TestServices.ReportAssertionFailure(
	testCase := _TestCase,
	message := _Message,
	sourceClassName := ClassName,
	defaultMessage := diagnostic
);
END_METHOD

END_FUNCTION_BLOCK

// ---- Assertions/TypedContexts/PointerAssertionContext.TcPOU
(*
SPDX-FileCopyrightText: © 2026 Oleksandr Tiutyk <trofimich@gmail.com>
SPDX-License-Identifier: MIT
License: https://opensource.org/license/mit
*)

(*!
<summary>Provides fluent assertions on a copied PVOID value.</summary>
<description>
Copies actual into persistent instance storage before the entry method returns; literals and expression
results therefore remain valid throughout the immediate chain. Owns no heap allocation or pointed-to resource.
The message prefixes every failure until the next preparation. Finish one chain before starting another on
the owning Assertions provider. Use only from the owning test callback on one task, without reentry.
Obtain this context from the owning provider; direct unprepared use is unsupported.
Expected arguments use the declared IEC type; ordinary compiler conversions happen before comparison.
This context does not depend on another assertion context.
Object metadata is available before preparation; inherited equality compares instance identity.
Copies the pointer value into a POINTER TO BYTE slot and never dereferences its target.
Equality compares addresses without generic conversion. Failed comparisons format the numeric addresses.
For interfaces and references, use ThatBool with the explicit null or validity predicate.
</description>
*)

{attribute 'no_explicit_call' := 'do not call this function block directly'}
FUNCTION_BLOCK PointerAssertionContext EXTENDS TOF_Core.Object
VAR_STAT
	{attribute 'hide'}
	_ClassName : STRING := __POUNAME();
END_VAR
VAR
	_Actual : POINTER TO BYTE;
	_TestCase : ITestCase;
	_Message : WSTRING(255);
END_VAR

(*!
<summary>Provides the implementation class name.</summary>
<description>
Borrowed read-only reference to compiler-initialized storage, valid throughout the instance lifetime.
Do not modify the returned reference; no ownership is transferred.
</description>
*)
{attribute 'monitoring' := 'call'}
PROPERTY ClassName : REFERENCE TO STRING
GET
ClassName REF= _ClassName;
END_GET
END_PROPERTY

(*!
<summary>Asserts that the copied pointer value is non-null.</summary>
<description>
Records failure without interrupting the callback; preserves the chain message.
</description>
*)
METHOD FINAL IsNotNull : REFERENCE TO PointerAssertionContext
IF _Actual = TOF_Core.Memory.NULL_ADDRESS THEN
	TestServices.ReportAssertionFailure(
		testCase := _TestCase,
		message := _Message,
		sourceClassName := ClassName,
		defaultMessage := "Expected: non-null object/pointer, but was null (0)"
	);
END_IF

IsNotNull REF= THIS^;
END_METHOD

(*!
<summary>Asserts that the copied pointer value is null.</summary>
<description>
Records failure without interrupting the callback; preserves the chain message.
</description>
*)
METHOD FINAL IsNull : REFERENCE TO PointerAssertionContext
IF _Actual <> TOF_Core.Memory.NULL_ADDRESS THEN
	TestServices.ReportAssertionFailure(
		testCase := _TestCase,
		message := _Message,
		sourceClassName := ClassName,
		defaultMessage := "Expected: null (0), but was non-zero address"
	);
END_IF

IsNull REF= THIS^;
END_METHOD

(*!
<summary>Provides the library namespace.</summary>
<description>
Borrowed read-only reference to the compiler-initialized namespace, valid throughout the instance lifetime.
Do not modify the returned reference; no ownership is transferred.
</description>
*)
{attribute 'monitoring' := 'call'}
PROPERTY NamespaceName : REFERENCE TO STRING
GET
NamespaceName REF= CurrentNamespace.Name;
END_GET
END_PROPERTY

(*!
<summary>Asserts inequality with the expected value.</summary>
<description>
Records failure without interrupting the callback; preserves the message for the rest of the chain.
</description>
<param name="expected">Expected value converted by the compiler to PVOID.</param>
*)
METHOD FINAL NotToBe : REFERENCE TO PointerAssertionContext
VAR_INPUT
	expected : PVOID;
END_VAR
IF _Actual = expected THEN
	failComparison(
		expected := expected,
		expectation := "Expected value not to be: "
	);
END_IF

NotToBe REF= THIS^;
END_METHOD

(*!
<summary>Copies the actual operand and replaces the chain-wide message.</summary>
<description>
Called by the owning Assertions provider after it verifies the running test case.
No pointer to this method's input storage is retained. The receiver is borrowed until the next preparation;
the owning provider keeps it alive throughout the immediate chain.
</description>
<param name="actual">Value copied into this context.</param>
<param name="testCase">Borrowed failure receiver for the immediate chain.</param>
<param name="message">Copied diagnostic prefix, including empty to clear the previous prefix.</param>
*)
METHOD INTERNAL FINAL Prepare
VAR_INPUT
	actual : PVOID;
	testCase : ITestCase;
	message : WSTRING(255);
END_VAR
_Actual := actual;
_TestCase := testCase;
_Message := message;
END_METHOD

(*!
<summary>Reports the byte size of this concrete instance.</summary>
<description>
Includes inline fields and nested instances, but excludes separately allocated payloads.
Obtaining the size does not transfer ownership or validate an arbitrary address.
</description>
*)
{attribute 'monitoring' := 'call'}
PROPERTY SelfSize : ULINT
GET
SelfSize := XSIZEOF(THIS^);
END_GET
END_PROPERTY

(*!
<summary>Asserts equality with the expected value.</summary>
<description>
Records failure without interrupting the callback; preserves the message for the rest of the chain.
</description>
<param name="expected">Expected value converted by the compiler to PVOID.</param>
*)
METHOD FINAL ToBe : REFERENCE TO PointerAssertionContext
VAR_INPUT
	expected : PVOID;
END_VAR
IF _Actual <> expected THEN
	failComparison(
		expected := expected,
		expectation := "Expected: "
	);
END_IF

ToBe REF= THIS^;
END_METHOD

(*!
<summary>Formats a failed typed predicate and reports it with the chain message.</summary>
<description>
Does not change operands or chain state. The receiver retains its first failure. Reporting exceptions
propagate to the enclosing test callback handler; an unprepared receiver is a configuration error.
</description>
<param name="expected">Typed expected operand used only for this diagnostic.</param>
<param name="expectation">Prefix identifying the failed predicate.</param>
*)
METHOD PRIVATE failComparison
VAR_INPUT
	expected : PVOID;
	expectation : WSTRING(40);
END_VAR
VAR
	actualText : WSTRING(255);
	expectedText : WSTRING(255);
	diagnostic : TOF_Core.ERROR_MESSAGE;
END_VAR
actualText := TO_WSTRING(TO_ULINT(_Actual));
expectedText := TO_WSTRING(TO_ULINT(expected));

diagnostic := TOF_Core.WideStrings.Concat255(
	expectation,
	expectedText,
	", but was: ",
	actualText
);

TestServices.ReportAssertionFailure(
	testCase := _TestCase,
	message := _Message,
	sourceClassName := ClassName,
	defaultMessage := diagnostic
);
END_METHOD

END_FUNCTION_BLOCK

// ---- TestElements/Groups/TestGroup.TcPOU
(*
SPDX-FileCopyrightText: © 2026 Oleksandr Tiutyk <trofimich@gmail.com>
SPDX-License-Identifier: MIT
License: https://opensource.org/license/mit
*)

(*!
<summary>Executes the fixed child array provided by a concrete group.</summary>
<description>
Descendants own persistent tests, nested groups and interface-array storage. Children returns the same valid
array throughout the group lifetime; callers must not modify its contents through the reference. Each child
is non-null, occurs once and has this group as its constructor-assigned Parent. Parent chains are acyclic.
All objects outlive the tree; no allocation ownership is transferred. Zero children form an empty group.
Reset validates the child reference, slots and parent chain once at the start of each run. Missing
array storage raises DataMemberNotSpecifiedException; null slots do likewise with an indexed member name.
Duplicates, a mismatched parent or a parent cycle raise StandardException before any direct child is called.
A descendant's validation or callback can still fail after earlier siblings have reset; no rollback is promised.
Execute drives one current child once and counts it once when finished. Groups add no synthetic test results
and have no scenario setup or teardown hooks. Use the entire tree in one task without reentry.
Do not mutate the child array or parent associations during the lifetime of the tree, or copy instances by value.
</description>
*)

{attribute 'no_explicit_call' := 'do not call this function block directly'}
FUNCTION_BLOCK ABSTRACT TestGroup
VAR_GENERIC CONSTANT
	//! <summary>Exact number of direct child slots; zero produces an empty array.</summary>
	{attribute 'hide'} 
	_ChildCount : TOF_Core.INT_LENGTH := 0;
END_VAR
EXTENDS TestElement IMPLEMENTS IParentTestElement
VAR
	{attribute 'hide'} 
	_CurrentChildIndex : TOF_Core.INT_LENGTH;
	
	{attribute 'hide'} 
	_TestCount : TOF_Core.DINT_LENGTH;
END_VAR

(*!
<summary>Reports the generic number of direct children.</summary>
*)

{attribute 'monitoring' := 'call'}
PROPERTY FINAL ChildCount : TOF_Core.INT_LENGTH
GET
ChildCount := _ChildCount;
END_GET
END_PROPERTY

(*!
<summary>Borrows the concrete group's persistent fixed array of tests and nested groups.</summary>
<description>
Return the same valid storage and unchanged child list for the group lifetime, including an empty array
when the generic count is zero. The getter must have no side effects. Callers may only read the reference.
Children are borrowed; each has this group as its fixed Parent and remains alive while the tree is used.
The base constructor never reads this property. Reset validates it before execution starts.
</description>
*)
{attribute 'monitoring' := 'call'}
PROPERTY ABSTRACT Children : REFERENCE TO ARRAY [0.._ChildCount - 1] OF ITestElement
GET
END_GET
END_PROPERTY

(*!
<summary>Advances one child of the validated fixed composition and counts it once on completion.</summary>
<description>
Requires a successful Reset before the first execution and every subsequent run, including after a failed Reset.
Uses the concrete group's Children reference without repeating topology validation.
External exceptions propagate to the runner and abort the run.
Neither Reset nor Execute changes parent associations.
</description>
*)
METHOD FINAL Execute
VAR
	childElements : REFERENCE TO ARRAY [0.._ChildCount - 1] OF ITestElement;
END_VAR
IF IsFinished THEN
	RETURN;
END_IF

childElements REF= THIS^.Children;

_State := TEST_ELEMENT_STATE.RUNNING;
_Duration := _Duration + TOF_Core.System.GetTaskCycleTime();

IF _CurrentChildIndex < _ChildCount THEN
	childElements[_CurrentChildIndex].Execute();

	IF childElements[_CurrentChildIndex].IsFinished THEN
		_PassedCount := _PassedCount + childElements[_CurrentChildIndex].PassedCount;
		_FailedCount := _FailedCount + childElements[_CurrentChildIndex].FailedCount;
		_SkippedCount := _SkippedCount + childElements[_CurrentChildIndex].SkippedCount;
		_CurrentChildIndex := _CurrentChildIndex + 1;
	END_IF

END_IF

IF _CurrentChildIndex >= _ChildCount THEN
	_State := TEST_ELEMENT_STATE.COMPLETED;
	_Reporter := 0;
END_IF
END_METHOD

(*!
<summary>Borrows one direct child in fixed execution order without changing the tree.</summary>
<description>
Checks storage before the index, including before the first Reset and after a failed Reset.
Missing storage or a null selected slot raises DataMemberNotSpecifiedException; an index outside
zero through ChildCount minus one raises ArgumentOutOfRangeException. No child callback is invoked.
The returned interface is borrowed for the child's lifetime. Use from the owning task without reentry;
this method does not repeat complete topology validation or authorize changes to the composition.
</description>
<param name="index">Zero-based position in the fixed direct-child array.</param>
*)
METHOD FINAL GetChildByIndex : ITestElement
VAR_INPUT
	index : TOF_Core.INT_LENGTH;
END_VAR
IF NOT __ISVALIDREF(Children) THEN
	TOF_Core.Exceptions.ThrowDataMemberNotSpecified(
		sourceNamespaceName := NamespaceName,
		sourceClassName := ClassName,
		sourcePOUName := __POUNAME(),
		sourcePosition := __POSITION(),
		dataMemberName := 'Children'
	);
END_IF

IF index < TOF_Core.SignedInt16.ZERO OR_ELSE index >= _ChildCount THEN
	TOF_Core.Exceptions.ThrowArgumentOutOfRange(
		sourceNamespaceName := NamespaceName,
		sourceClassName := ClassName,
		sourcePOUName := __POUNAME(),
		sourcePosition := __POSITION(),
		argumentName := 'index',
		argumentValue := index
	);
END_IF

IF Children[index] = 0 THEN
	TOF_Core.Exceptions.ThrowDataMemberNotSpecified(
		sourceNamespaceName := NamespaceName,
		sourceClassName := ClassName,
		sourcePOUName := __POUNAME(),
		sourcePosition := __POSITION(),
		dataMemberName := TOF_Core.Strings.Concat255('Children[', TO_STRING(index), ']')
	);
END_IF

GetChildByIndex := Children[index];
END_METHOD

//! <summary>Sums the leaf counts of the group's direct children.</summary>
METHOD PRIVATE getTestCount : TOF_Core.DINT_LENGTH
VAR
	// An empty group gives the FOR loop an upper bound of -1.
	i : INT;
END_VAR
IF NOT __ISVALIDREF(Children) THEN
	RETURN;
END_IF

FOR i := 0 TO _ChildCount - 1 DO
	getTestCount := getTestCount + Children[i].TestCount;
END_FOR
END_METHOD

(*!
<summary>Clears observations and recursively resets descendant-specific state.</summary>
<description>
Does not run teardown or release user resources. Call only at the lifecycle boundaries in ITestElement.
The reporter is borrowed until completion; no locks or cross-task transfer are provided.
Validation or a child Reset exception propagates and can leave a partially reset tree; the runner aborts startup.
</description>
*)
METHOD FINAL Reset
VAR_INPUT
	reporter : ITestReporter;
END_VAR
VAR
	self : ITestElement;
	slowAncestor : ITestElement;
	fastAncestor : ITestElement;
	childParent : ITestElement;

	i : INT;
	j : INT;
	
	errorMessage : TOF_Core.ERROR_MESSAGE;
END_VAR
SUPER^.Reset(reporter := reporter);

IF NOT __ISVALIDREF(Children) THEN
	TOF_Core.Exceptions.ThrowDataMemberNotSpecified(
		sourceNamespaceName := NamespaceName,
		sourceClassName := ClassName,
		sourcePOUName := __POUNAME(),
		sourcePosition := __POSITION(),
		dataMemberName := 'Children'
	);
END_IF

self := THIS^;
slowAncestor := self;
fastAncestor := self;

// Traverse the fixed parent chain at two speeds to detect cycles without allocation or recursion.
WHILE fastAncestor <> 0 DO
	fastAncestor := fastAncestor.Parent;

	IF fastAncestor = 0 THEN
		EXIT;
	END_IF

	fastAncestor := fastAncestor.Parent;
	slowAncestor := slowAncestor.Parent;

	IF fastAncestor <> 0 AND_THEN fastAncestor = slowAncestor THEN
		TOF_Core.Exceptions.ThrowStandard(
			sourceNamespaceName := NamespaceName,
			sourceClassName := ClassName,
			sourcePOUName := __POUNAME(),
			sourcePosition := __POSITION(),
			message := "The assigned parent chain contains a cycle"
		);
	END_IF
END_WHILE

FOR i := 0 TO _ChildCount - 1 DO
	IF Children[i] = 0 THEN
		TOF_Core.Exceptions.ThrowDataMemberNotSpecified(
			sourceNamespaceName := NamespaceName,
			sourceClassName := ClassName,
			sourcePOUName := __POUNAME(),
			sourcePosition := __POSITION(),
			dataMemberName := TOF_Core.Strings.Concat255('Children[', TO_STRING(i), ']')
		);
	END_IF

	childParent := Children[i].Parent;

	IF childParent <> self THEN
		errorMessage := TOF_Core.WideStrings.Concat255("A child '", Children[i].Name, "' has a different constructor-assigned parent"); 
		
		TOF_Core.Exceptions.ThrowStandard(
			sourceNamespaceName := NamespaceName,
			sourceClassName := ClassName,
			sourcePOUName := __POUNAME(),
			sourcePosition := __POSITION(),
			message := errorMessage
		);
	END_IF

	FOR j := 0 TO i - 1 DO
		IF Children[i] = Children[j] THEN
			errorMessage := TOF_Core.WideStrings.Concat255("A child '", Children[i].Name, "' occupies more than one slot"); 
			
			TOF_Core.Exceptions.ThrowStandard(
				sourceNamespaceName := NamespaceName,
				sourceClassName := ClassName,
				sourcePOUName := __POUNAME(),
				sourcePosition := __POSITION(),
				message := errorMessage
			);
		END_IF
	END_FOR
END_FOR

_CurrentChildIndex := 0;

FOR i := 0 TO _ChildCount - 1 DO
	Children[i].Reset(reporter := _Reporter);
END_FOR
END_METHOD

(*!
<summary>Sums the configured leaf counts of the direct children.</summary>
<description>
Requires a valid, acyclic subtree. Traverses nested groups through their getters using the current task stack.
An empty group returns zero. Missing child storage or a null slot in a nonempty group raises
DataMemberNotSpecifiedException. Child getter exceptions propagate and the tree state is unchanged.
</description>
*)
{attribute 'monitoring' := 'call'}
PROPERTY FINAL TestCount : TOF_Core.DINT_LENGTH
GET
IF _TestCount = 0 THEN
	_TestCount := getTestCount();
END_IF

TestCount := _TestCount;
END_GET
END_PROPERTY

END_FUNCTION_BLOCK

// ---- Reporting/AdsLogReporter.TcPOU
(*
SPDX-FileCopyrightText: © 2026 Oleksandr Tiutyk <trofimich@gmail.com>
SPDX-License-Identifier: MIT
License: https://opensource.org/license/mit
*)

(*!
<summary>Writes run summaries and leaf failures to the ADS log.</summary>
<description>
Use in one task without reentry. The ADS backend has no established concurrent-call guarantee, even for
separate reporter instances. For multiple tasks use per-task in-memory reports or a synchronized backend.
Each callback submits at most one record. The ADS completion record includes counts and the first failed leaf name.
LastRunSummary includes the first failed leaf name and a bounded
version of its diagnostic. The summary and failed log writes are observable after the run. A failed
write does not change the test outcome. Individual ADS failure records are capped at 200 wide characters.
ReportRunStart clears all observations before attempting the start message.
</description>
*)

{attribute 'no_explicit_call' := 'do not call this function block directly'}
FUNCTION_BLOCK AdsLogReporter EXTENDS TOF_Core.Object IMPLEMENTS ITestReporter
VAR_STAT
	_ClassName : STRING := __POUNAME();
END_VAR
VAR
	_AdsLogger : TOF_Core.AdsLogger;
	_FirstFailureName : WSTRING;
	_FirstFailureDiagnostic : WSTRING(255);
	_LastRunSummary : TOF_Core.ERROR_MESSAGE;
	_FailedLogWriteCount : UDINT;
	_LastLogFailureMessage : TOF_Core.ERROR_MESSAGE;
END_VAR

(*!
<summary>Provides the implementation class name.</summary>
*)
{attribute 'monitoring' := 'call'}
PROPERTY ClassName : REFERENCE TO STRING
GET
ClassName REF= _ClassName;
END_GET
END_PROPERTY

(*!
<summary>Counts start, result and summary writes for which TryLogMessage returned FALSE.</summary>
<description>The count resets at ReportRunStart. A successful write does not confirm display in XAE.</description>
*)
{attribute 'monitoring' := 'call'}
PROPERTY FailedLogWriteCount : UDINT
GET
FailedLogWriteCount := _FailedLogWriteCount;
END_GET
END_PROPERTY

(*!
<summary>Borrows the last message whose ADS logger call returned FALSE.</summary>
<description>Empty until a write fails in the current run. Callers must not modify the returned storage.</description>
*)
{attribute 'monitoring' := 'call'}
PROPERTY LastLogFailureMessage : REFERENCE TO TOF_Core.ERROR_MESSAGE
GET
LastLogFailureMessage REF= _LastLogFailureMessage;
END_GET
END_PROPERTY

(*!
<summary>Borrows the summary created at ReportRunEnd regardless of its ADS write status.</summary>
<description>Empty after ReportRunStart until ReportRunEnd. Callers must not modify the returned storage.</description>
*)
{attribute 'monitoring' := 'call'}
PROPERTY LastRunSummary : REFERENCE TO TOF_Core.ERROR_MESSAGE
GET
LastRunSummary REF= _LastRunSummary;
END_GET
END_PROPERTY

(*!
<summary>Submits one ADS message and records a FALSE result from the logger.</summary>
<description>The count saturates at the largest UDINT. The copied text remains available until the next start.</description>
*)
METHOD PRIVATE logMessage
VAR_INPUT
	category : TOF_Core.LOG_CATEGORY;
END_VAR
VAR_IN_OUT CONSTANT
	message : TOF_Core.ERROR_MESSAGE;
END_VAR
IF TryWriteMessage(category := category, message := message) THEN
	RETURN;
END_IF

IF _FailedLogWriteCount < TOF_Core.UnsignedInt32.MAX_VALUE THEN
	_FailedLogWriteCount := _FailedLogWriteCount + 1;
END_IF

_LastLogFailureMessage := message;
END_METHOD

(*!
<summary>Provides the library namespace.</summary>
*)
{attribute 'monitoring' := 'call'}
PROPERTY NamespaceName : REFERENCE TO STRING
GET
NamespaceName REF= CurrentNamespace.Name;
END_GET
END_PROPERTY

(*!
<summary>Logs leaf counts and the first failed leaf name and retains its diagnostic for online inspection.</summary>
<description>The retained summary also includes a bounded first-failure diagnostic and survives a rejected ADS write.</description>
*)
METHOD ReportRunEnd
VAR_INPUT
	totalTests : TOF_Core.DINT_LENGTH;
	passedTests : TOF_Core.DINT_LENGTH;
	failedTests : TOF_Core.DINT_LENGTH;
	skippedTests : TOF_Core.DINT_LENGTH;
	duration : TIME;
END_VAR
VAR
	logSummary : WSTRING(255);
	logRecord : TOF_Core.ERROR_MESSAGE;
	summary : WSTRING(255);
END_VAR
summary := TOF_Core.WideStrings.Concat255(
	"[TOF_Testing] Finished: ", TO_WSTRING(passedTests), " passed, ",
	TO_WSTRING(failedTests), " failed, ", TO_WSTRING(skippedTests), " skipped"
);

logSummary := summary;

IF failedTests > 0 AND_THEN _FirstFailureDiagnostic <> "" THEN
	TOF_Core.WideStrings.AppendFit255(logSummary, " | First failed test: ", _FirstFailureName);
	TOF_Core.WideStrings.AppendFit255(summary, " | First failure: ", _FirstFailureDiagnostic);
END_IF

_LastRunSummary := summary;
logRecord := logSummary;
logMessage(category := TOF_Core.LOG_CATEGORY.INFORMATION, message := logRecord);
END_METHOD

(*!
<summary>Resets per-run observations and logs the number of configured leaf tests.</summary>
<description>A failed start-message write counts toward the new run.</description>
*)
METHOD ReportRunStart
VAR_INPUT
	testCount : TOF_Core.DINT_LENGTH;
END_VAR
VAR
	diagnostic : TOF_Core.ERROR_MESSAGE;
END_VAR
_FirstFailureName := "";
_FirstFailureDiagnostic := "";
_LastRunSummary := "";
_FailedLogWriteCount := 0;
_LastLogFailureMessage := "";

diagnostic := TOF_Core.WideStrings.Concat255(
	"[TOF_Testing] Starting ", TO_WSTRING(testCount), " tests"
);

logMessage(category := TOF_Core.LOG_CATEGORY.INFORMATION, message := diagnostic);
END_METHOD

(*!
<summary>Logs a failed leaf with its group path and caches the first failure for the summary.</summary>
<description>
The individual ADS record uses up to 200 wide characters to leave room below the native ADS text limit.
The retained summary includes the leaf name and the beginning of its diagnostic.
</description>
<param name="testName">Individual name bounded to 80 wide characters, matching INamed.</param>
*)
METHOD ReportTestCaseResult
VAR_INPUT
	groupPath : WSTRING(255);
	testName : WSTRING;
	outcome : TEST_OUTCOME;
	duration : TIME;
END_VAR
VAR_IN_OUT CONSTANT
	message : TOF_Core.ERROR_MESSAGE;
END_VAR
VAR
	shortDiagnostic : WSTRING(200);
	diagnostic : TOF_Core.ERROR_MESSAGE;
END_VAR
IF outcome <> TEST_OUTCOME.PASSED
	AND_THEN outcome <> TEST_OUTCOME.FAILED
	AND_THEN outcome <> TEST_OUTCOME.SKIPPED
THEN
	TOF_Core.Exceptions.ThrowArgumentValueNotSupported(
		sourceNamespaceName := NamespaceName,
		sourceClassName := ClassName,
		sourcePOUName := __POUNAME(),
		sourcePosition := __POSITION(),
		argumentName := 'outcome',
		argumentValue := outcome
	);
END_IF

IF outcome <> TEST_OUTCOME.FAILED THEN
	RETURN;
END_IF

IF _FirstFailureDiagnostic = "" THEN
	_FirstFailureName := testName;

	IF _FirstFailureName = "" THEN
		_FirstFailureName := "<unnamed>";
	END_IF

	_FirstFailureDiagnostic := TOF_Core.WideStrings.Concat255(_FirstFailureName, ": ");
	TOF_Core.WideStrings.AppendFit(targetString := _FirstFailureDiagnostic, sourceString := message);
END_IF

shortDiagnostic := "[TOF_Testing] ";

IF groupPath <> "" THEN
	TOF_Core.WideStrings.AppendFit255(shortDiagnostic, groupPath, "/");
END_IF

TOF_Core.WideStrings.AppendFit255(shortDiagnostic, testName, ": ");
TOF_Core.WideStrings.AppendFit(targetString := shortDiagnostic, sourceString := message);
diagnostic := shortDiagnostic;

logMessage(category := TOF_Core.LOG_CATEGORY.ERROR, message := diagnostic);
END_METHOD

(*!
<summary>Reports instance storage without separately allocated payloads.</summary>
*)
{attribute 'monitoring' := 'call'}
PROPERTY SelfSize : ULINT
GET
SelfSize := XSIZEOF(THIS^);
END_GET
END_PROPERTY

(*!
<summary>Submits one message to the ADS backend and reports whether the logger accepted it.</summary>
<description>
An override may replace the backend. It must return FALSE on rejection and must not raise an exception,
retry the write, or retain the borrowed message. TRUE does not confirm display in XAE.
</description>
*)
METHOD PROTECTED TryWriteMessage : BOOL
VAR_INPUT
	category : TOF_Core.LOG_CATEGORY;
END_VAR
VAR_IN_OUT CONSTANT
	message : TOF_Core.ERROR_MESSAGE;
END_VAR
TryWriteMessage := _AdsLogger.TryLogMessage(category := category, message := message);
END_METHOD

END_FUNCTION_BLOCK

// ---- Reporting/JUnitXmlReporter.TcPOU
(*
SPDX-FileCopyrightText: © 2026 Oleksandr Tiutyk <trofimich@gmail.com>
SPDX-License-Identifier: MIT
License: https://opensource.org/license/mit
*)

(*!
<summary>Builds an in-memory JUnit report with one testcase per leaf.</summary>
<description>
One flat testsuite contains all leaves; testcase classname preserves the slash-separated group path.
Wide names and diagnostics are escaped as ASCII XML character references, including surrogate pairs.
XML 1.0 disallowed control characters, isolated surrogates and U+FFFE/U+FFFF are replaced by U+FFFD;
tab, line feed and carriage return are emitted as references to preserve attribute whitespace.
Use a separate instance and buffer for each runner task without reentry. Read ContentLength bytes from
ContentAddress only after IsReady and before reset or the next run. Buffer growth invalidates old addresses.
The reporter owns its dynamic buffer; never copy it by value. Callback exceptions can leave incomplete XML.
</description>
*)

{attribute 'no_explicit_call' := 'do not call this function block directly'}
FUNCTION_BLOCK JUnitXmlReporter EXTENDS TOF_Core.Object IMPLEMENTS ITestReporter
VAR CONSTANT
	//! <summary>First and last UTF-16 high-surrogate code units; subtract the first to recover ten payload bits.</summary>
	HIGH_SURROGATE_FIRST : UDINT := 16#D800;
	//! <summary>Last UTF-16 high-surrogate code unit accepted as the first part of a pair.</summary>
	HIGH_SURROGATE_LAST : UDINT := 16#DBFF;
	//! <summary>First and last UTF-16 low-surrogate code units; subtract the first to recover ten payload bits.</summary>
	LOW_SURROGATE_FIRST : UDINT := 16#DC00;
	//! <summary>Last UTF-16 low-surrogate code unit; isolated surrogates through this value are invalid scalars.</summary>
	LOW_SURROGATE_LAST : UDINT := 16#DFFF;
	//! <summary>Base scalar value added when decoding a supplementary UTF-16 surrogate pair.</summary>
	SUPPLEMENTARY_FIRST : UDINT := 16#10000;
	//! <summary>Multiplier that moves a high surrogate's ten payload bits above the low payload.</summary>
	SURROGATE_PAYLOAD_BASE : UDINT := 1024;
	//! <summary>Printable ASCII boundaries; these scalars are emitted as bytes instead of decimal XML references.</summary>
	PRINTABLE_ASCII_FIRST : UDINT := 32;
	//! <summary>Last ASCII scalar emitted directly as a byte instead of a decimal XML reference.</summary>
	PRINTABLE_ASCII_LAST : UDINT := 126;
END_VAR
VAR_STAT
	_ClassName : STRING := __POUNAME();
END_VAR
VAR
	_Buffer : TOF_Core.StringBuilder;
	_IsReady : BOOL;
END_VAR

//! <summary>Escapes UTF-16 input and replaces isolated surrogates and forbidden XML characters.</summary>
METHOD PRIVATE appendEscapedText
VAR_IN_OUT CONSTANT
	text : WSTRING;
END_VAR
VAR
	charLength : UDINT;
	i : UDINT;
	wordPointer : POINTER TO WORD;
	codePoint : UDINT;
END_VAR
charLength := TOF_Core.WideStrings.GetLength(value := text);
wordPointer := ADR(text);

WHILE i < charLength DO
	codePoint := wordPointer[i];
	i := i + 1;

	IF codePoint >= HIGH_SURROGATE_FIRST AND_THEN codePoint <= HIGH_SURROGATE_LAST AND_THEN i < charLength
		AND_THEN wordPointer[i] >= LOW_SURROGATE_FIRST AND_THEN wordPointer[i] <= LOW_SURROGATE_LAST
	THEN
		// UTF-16 uses high D800..DBFF and low DC00..DFFF surrogates. Subtract their bases to obtain
		// ten-bit payloads; shift the high payload by ten bits and add the supplementary-plane base.
		codePoint := SUPPLEMENTARY_FIRST + (codePoint - HIGH_SURROGATE_FIRST) * SURROGATE_PAYLOAD_BASE
			+ (wordPointer[i] - LOW_SURROGATE_FIRST);
		i := i + 1;
	END_IF

	appendXmlCharacter(codePoint := codePoint);
END_WHILE
END_METHOD

(*!
<summary>Appends a scalar as printable ASCII or an XML decimal character reference.</summary>
<description>Explicitly terminates the single-byte temporary before the buffer reads it.</description>
*)
METHOD PRIVATE appendXmlCharacter
VAR_INPUT
	codePoint : UDINT;
END_VAR
VAR
	character : STRING(1);
	referenceText : STRING(255);
END_VAR
// XML 1.0 permits only TAB/LF/CR below U+0020 and excludes surrogates and U+FFFE/U+FFFF.
CASE codePoint OF
	0..8, 11, 12, 14..31, 16#D800..16#DFFF, 16#FFFE, 16#FFFF:
		_Buffer.AppendString(value := '&#65533;');
	34:
		_Buffer.AppendString(value := '&quot;');
	38:
		_Buffer.AppendString(value := '&amp;');
	39:
		_Buffer.AppendString(value := '&apos;');
	60:
		_Buffer.AppendString(value := '&lt;');
	62:
		_Buffer.AppendString(value := '&gt;');
ELSE
	IF codePoint >= PRINTABLE_ASCII_FIRST AND_THEN codePoint <= PRINTABLE_ASCII_LAST THEN
		character[0] := TO_BYTE(codePoint);
		character[1] := TO_BYTE(TOF_Core.UnsignedInt8.MIN_VALUE);
		_Buffer.AppendString(value := character);
	ELSE
		referenceText := TOF_Core.Strings.Concat255('&#', TO_STRING(codePoint), ';');
		_Buffer.AppendString(value := referenceText);
	END_IF
END_CASE
END_METHOD

(*!
<summary>Provides the implementation class name.</summary>
*)
{attribute 'monitoring' := 'call'}
PROPERTY ClassName : REFERENCE TO STRING
GET
ClassName REF= _ClassName;
END_GET
END_PROPERTY

(*!
<summary>Borrows the current XML buffer address.</summary>
*)
{attribute 'monitoring' := 'call'}
PROPERTY ContentAddress : POINTER TO STRING
GET
ContentAddress := _Buffer.StringAddress;
END_GET
END_PROPERTY

(*!
<summary>Reports the ASCII byte count excluding the terminating zero.</summary>
*)
{attribute 'monitoring' := 'call'}
PROPERTY ContentLength : UDINT
GET
ContentLength := _Buffer.StringLength;
END_GET
END_PROPERTY

(*!
<summary>Reports whether ReportRunEnd completed the XML document.</summary>
*)
{attribute 'monitoring' := 'call'}
PROPERTY IsReady : BOOL
GET
IsReady := _IsReady;
END_GET
END_PROPERTY

(*!
<summary>Provides the library namespace.</summary>
*)
{attribute 'monitoring' := 'call'}
PROPERTY NamespaceName : REFERENCE TO STRING
GET
NamespaceName REF= CurrentNamespace.Name;
END_GET
END_PROPERTY

(*!
<summary>Closes the JUnit container and makes its buffer available to readers.</summary>
*)
METHOD ReportRunEnd
VAR_INPUT
	totalTests : TOF_Core.DINT_LENGTH;
	passedTests : TOF_Core.DINT_LENGTH;
	failedTests : TOF_Core.DINT_LENGTH;
	skippedTests : TOF_Core.DINT_LENGTH;
	duration : TIME;
END_VAR
_Buffer.AppendString(value := '  </testsuite>$R$N</testsuites>$R$N');
_IsReady := TRUE;
END_METHOD

(*!
<summary>Clears previous output and opens the flat JUnit container.</summary>
<param name="testCount">Planned leaf count. The XML summary uses actual results supplied at run end.</param>
*)
METHOD ReportRunStart
VAR_INPUT
	testCount : TOF_Core.DINT_LENGTH;
END_VAR
_Buffer.Clear(releaseMemory := FALSE);
_IsReady := FALSE;
_Buffer.AppendString(value := '<?xml version="1.0" encoding="UTF-8"?>$R$N');
_Buffer.AppendString(value := '<testsuites>$R$N  <testsuite name="OpenFramework">$R$N');
END_METHOD

(*!
<summary>Appends a terminal leaf result with its group path as classname.</summary>
<param name="testName">Individual name bounded to 80 wide characters, matching INamed.</param>
*)
METHOD ReportTestCaseResult
VAR_INPUT
	groupPath : WSTRING(255);
	testName : WSTRING;
	outcome : TEST_OUTCOME;
	duration : TIME;
END_VAR
VAR_IN_OUT CONSTANT
	message : TOF_Core.ERROR_MESSAGE;
END_VAR
VAR
	milliseconds : UDINT;
	timeAttribute : STRING(255);
END_VAR
IF outcome <> TEST_OUTCOME.PASSED
	AND_THEN outcome <> TEST_OUTCOME.FAILED
	AND_THEN outcome <> TEST_OUTCOME.SKIPPED
THEN
	TOF_Core.Exceptions.ThrowArgumentValueNotSupported(
		sourceNamespaceName := NamespaceName,
		sourceClassName := ClassName,
		sourcePOUName := __POUNAME(),
		sourcePosition := __POSITION(),
		argumentName := 'outcome',
		argumentValue := outcome
	);
END_IF

_Buffer.AppendString(value := '    <testcase name="');
appendEscapedText(text := testName);
_Buffer.AppendString(value := '" classname="');
appendEscapedText(text := groupPath);
milliseconds := TO_UDINT(duration);
timeAttribute := TOF_Core.Strings.Concat255(
	'" time="',
	TO_STRING(milliseconds / 1000),
	'.',
	TO_STRING(milliseconds / 100 MOD 10),
	TO_STRING(milliseconds / 10 MOD 10),
	TO_STRING(milliseconds MOD 10),
	'"'
);
_Buffer.AppendString(value := timeAttribute);

IF outcome = TEST_OUTCOME.FAILED THEN
	_Buffer.AppendString(value := '>$R$N');
	_Buffer.AppendString(value := '      <failure message="');
	appendEscapedText(text := message);
	_Buffer.AppendString(value := '" type="AssertionFailure">');
	appendEscapedText(text := message);
	_Buffer.AppendString(value := '</failure>$R$N');
	_Buffer.AppendString(value := '    </testcase>$R$N');
ELSIF outcome = TEST_OUTCOME.SKIPPED THEN
	_Buffer.AppendString(value := '>$R$N');
	_Buffer.AppendString(value := '      <skipped />$R$N');
	_Buffer.AppendString(value := '    </testcase>$R$N');
ELSE
	_Buffer.AppendString(value := ' />$R$N');
END_IF
END_METHOD

(*!
<summary>Releases the XML buffer outside an active run; existing reader addresses become invalid.</summary>
*)
METHOD FINAL Reset
_Buffer.Clear(releaseMemory := TRUE);

_IsReady := FALSE;
END_METHOD

(*!
<summary>Reports instance storage without separately allocated payloads.</summary>
*)
{attribute 'monitoring' := 'call'}
PROPERTY SelfSize : ULINT
GET
SelfSize := XSIZEOF(THIS^);
END_GET
END_PROPERTY

END_FUNCTION_BLOCK

// ---- Runner/TestRunner.TcPOU
(*
SPDX-FileCopyrightText: © 2026 Oleksandr Tiutyk <trofimich@gmail.com>
SPDX-License-Identifier: MIT
License: https://opensource.org/license/mit
*)

(*!
<summary>Runs a fixed tree of individual tests and nested groups in its owning PLC task.</summary>
<description>
Concrete descendants own their persistent root tests, groups and interface-array storage and provide Children.
Call Execute once per PLC cycle until IsFinished. Each run validates roots in STARTING before any direct Reset
or report callback. Missing storage or null slots raise DataMemberNotSpecifiedException; duplicates, running
or group-owned roots raise StandardException. Execute catches these failures and exposes an aborted run.
Children returns the same valid storage and unchanged list throughout the runner lifetime; do not mutate it.
After startup the runner advances at most one leaf body per call without repeating topology checks.
AllPassed is meaningful only after IsFinished. Roots are constructed with parent := 0; Parent is the fixed association with a group.
Register each root instance with one runner only and keep the tree stable. This is a caller
precondition: no parent marker or registry detects sharing roots between runners. Empty runs pass with zero tests.
ExitCode is the failed leaf count, or -1 for a startup failure or an aborted
external callback. An aborted callback is never retried; partial counts and report output are possible.
Before Reset of an externally aborted tree, make its user resources safe; Reset does not provide cancellation.
Use one task without reentry per runner, tree and reporter. Other tasks need disjoint instances and buffers.
Mutable tested resources and custom callbacks also require task isolation or their own synchronization.
The default ADS backend has no established concurrent-call guarantee; use a separate JUnitXmlReporter per task
for independent in-memory reporting, or a reporter backed by a synchronized logging service.
Execute enforces terminal OOM outside recoverable catches. Standalone execution uses cleanupTaskMemory := TRUE
(the default) to clean the current task after the last consumer of transient exceptions. Under AutomationRunner
or any other host that performs this cleanup at the task boundary, pass cleanupTaskMemory := FALSE.
This runner borrows its children and reporter; never copy it by value or delete dependencies while attached.
</description>
*)

{attribute 'no_explicit_call' := 'do not call this function block directly'}
FUNCTION_BLOCK ABSTRACT TestRunner
VAR_GENERIC CONSTANT
	//! <summary>Exact number of root test or group slots.</summary>
	_ChildCount : TOF_Core.INT_LENGTH := 0;
END_VAR
EXTENDS TOF_Core.Object
VAR_OUTPUT
	IsFinished : BOOL;
	AllPassed : BOOL;
	ExitCode : DINT;
	//! <summary>Runtime exception code for startup or external callback failure when ExitCode is -1.</summary>
	CallbackException : __SYSTEM.ExceptionCode;
	//! <summary>Copied stage and exception diagnostic for the aborted run; empty after Reset.</summary>
	CallbackMessage : TOF_Core.ERROR_MESSAGE;
	TotalTests : TOF_Core.DINT_LENGTH;
	PassedTests : TOF_Core.DINT_LENGTH;
	FailedTests : TOF_Core.DINT_LENGTH;
	SkippedTests : TOF_Core.DINT_LENGTH;
	TotalDuration : TIME;
END_VAR
VAR
	_CurrentChildIndex : TOF_Core.INT_LENGTH;
	_Duration : LTIME;
	_Reporter : ITestReporter;
	_DefaultAdsReporter : AdsLogReporter;
	_State : TEST_RUN_PHASE;
END_VAR

(*!
<summary>Reports the generic number of direct children.</summary>
*)

{attribute 'monitoring' := 'call'}
PROPERTY FINAL ChildCount : TOF_Core.INT_LENGTH
GET
ChildCount := _ChildCount;
END_GET
END_PROPERTY

(*!
<summary>Borrows the concrete runner's unchanged persistent array of parentless roots.</summary>
<description>
Return the same valid storage and unchanged list for the runner lifetime, including an empty array when N is zero.
The getter has no side effects. Callers may only read the reference; each root belongs to this runner alone.
The concrete descendant owns persistent roots and array storage. Roots use parent := 0 and outlive every run.
The base constructor never reads this property. Validation starts in Execute after construction.
</description>
*)
{attribute 'monitoring' := 'call'}
PROPERTY ABSTRACT Children : REFERENCE TO ARRAY [0.._ChildCount - 1] OF ITestElement
GET
END_GET
END_PROPERTY

(*!
<summary>Drives one root cycle and enforces the terminal allocation latch at the task boundary.</summary>
<description>
Catches startup validation and external callback failures to abort with ExitCode -1, then raises terminal OOM
outside the recoverable catch regardless of cleanupTaskMemory.
With cleanupTaskMemory TRUE, cleans all registered auto-disposed objects and the exception payload of the current
PLC task before returning, not only objects created by this runner. Borrowed references to those objects become
invalid; call after the last consumer of transient exceptions in the task cycle.
With cleanupTaskMemory FALSE, the host must call DynamicMemoryManager.RaiseIfAllocationFailed outside recoverable
handlers, then DynamicMemoryManager.CleanupMemory after all transient-exception consumers in each task cycle.
For multiple runners in one task, pass FALSE to each and let the host provide the shared task boundary.
</description>
<param name="cleanupTaskMemory">
TRUE by default for standalone execution. Pass FALSE under AutomationRunner or any other host that performs
current-task memory cleanup after all transient-exception consumers.
</param>
*)
METHOD FINAL Execute
VAR_INPUT
	cleanupTaskMemory : BOOL := TRUE;
END_VAR
VAR
	exceptionCode : __SYSTEM.ExceptionCode;
END_VAR
__TRY
	executeCycle();
__CATCH(exceptionCode)
	CallbackException := exceptionCode;
	CallbackMessage := TestServices.FormatCaughtException(
		exceptionCode := exceptionCode,
		stage := TO_STRING(_State),
		catchPointPOUName := __POUNAME(),
		catchPointPosition := __POSITION()
	);
	AllPassed := FALSE;
	ExitCode := -1;
	IsFinished := TRUE;
	_State := TEST_RUN_PHASE.COMPLETED;
__ENDTRY

TOF_Core.DynamicMemoryManager.RaiseIfAllocationFailed();

IF cleanupTaskMemory THEN
	TOF_Core.DynamicMemoryManager.CleanupMemory();
END_IF
END_METHOD

(*!
<summary>Advances one direct child and synchronously delivers run-level reporter callbacks.</summary>
<description>
Validates the fixed roots once in STARTING before direct Reset or reporting; callbacks may partially reset the tree.
After all roots reset successfully, reports the summed leaf count, including tests that may later be skipped.
</description>
*)
METHOD PRIVATE executeCycle
VAR
	activeReporter : ITestReporter;
	
	testCount : TOF_Core.DINT_LENGTH;
	
	i : INT;
END_VAR
IF _Reporter <> 0 THEN
	activeReporter := _Reporter;
ELSE
	activeReporter := _DefaultAdsReporter;
END_IF

CASE _State OF
	TEST_RUN_PHASE.STARTING:
		validateChildren(rejectRunningChildren := TRUE);

		_CurrentChildIndex := 0;
		_Duration := LTIME#0NS;

		FOR i := 0 TO _ChildCount - 1 DO
			Children[i].Reset(reporter := activeReporter);
		END_FOR

		testCount := 0;

		FOR i := 0 TO _ChildCount - 1 DO
			testCount := testCount + Children[i].TestCount;
		END_FOR

		activeReporter.ReportRunStart(testCount := testCount);
		
		_State := TEST_RUN_PHASE.RUNNING_ELEMENTS;

	TEST_RUN_PHASE.RUNNING_ELEMENTS:
		_Duration := _Duration + TOF_Core.System.GetTaskCycleTime();

		IF _CurrentChildIndex < _ChildCount THEN
			Children[_CurrentChildIndex].Execute();

			IF Children[_CurrentChildIndex].IsFinished THEN
				PassedTests := PassedTests + Children[_CurrentChildIndex].PassedCount;
				FailedTests := FailedTests + Children[_CurrentChildIndex].FailedCount;
				SkippedTests := SkippedTests + Children[_CurrentChildIndex].SkippedCount;
				
				_CurrentChildIndex := _CurrentChildIndex + 1;
			END_IF

		END_IF

		TotalTests := PassedTests + FailedTests + SkippedTests;
		TotalDuration := TO_TIME(_Duration);

		IF _CurrentChildIndex >= _ChildCount THEN
			_State := TEST_RUN_PHASE.REPORTING_TOTALS;
		END_IF

	TEST_RUN_PHASE.REPORTING_TOTALS:
		activeReporter.ReportRunEnd(
			totalTests := TotalTests,
			passedTests := PassedTests,
			failedTests := FailedTests,
			skippedTests := SkippedTests,
			duration := TotalDuration
		);
		
		AllPassed := (FailedTests = TOF_Core.SignedInt32.ZERO);
		ExitCode := TO_DINT(FailedTests);
		IsFinished := TRUE;
		
		_State := TEST_RUN_PHASE.COMPLETED;

	TEST_RUN_PHASE.COMPLETED:
		;
END_CASE
END_METHOD

(*!
<summary>Gets or configures the borrowed reporter; zero selects the ADS reporter.</summary>
<description>
Keep the same reporter alive throughout the run. Mutation during execution raises StandardException;
the failure concerns the active state rather than the requested reporter value.
</description>
*)
{attribute 'monitoring' := 'call'}
PROPERTY Reporter : ITestReporter
GET
Reporter := _Reporter;
END_GET
SET
IF _State = TEST_RUN_PHASE.RUNNING_ELEMENTS OR_ELSE _State = TEST_RUN_PHASE.REPORTING_TOTALS THEN
	TOF_Core.Exceptions.ThrowStandard(
		sourceNamespaceName := NamespaceName,
		sourceClassName := ClassName,
		sourcePOUName := __POUNAME(),
		sourcePosition := __POSITION(),
		message := "Cannot change the active reporter"
	);
END_IF

_Reporter := Reporter;
END_SET
END_PROPERTY

(*!
<summary>Rearms a completed or not-yet-started runner; calls during a normal run are ignored.</summary>
<description>
The next Execute resets the tree. After an external callback abort the caller must first recover any
user resources not covered by scenario teardown. After abort, Reset validates root storage and topology and recursively
resets the same tree immediately, without setup, body, teardown or reporter callbacks.
Running roots are allowed during abort recovery. A validation failure calls no child and retains the aborted observations.
Custom element Reset callbacks can throw; runner observations remain aborted and recovery can be retried.
Other tree resets remain deferred until Execute. Reset does not clear terminal allocation failure.
</description>
*)
METHOD FINAL Reset
VAR
	i : INT;
END_VAR
IF _State = TEST_RUN_PHASE.RUNNING_ELEMENTS OR_ELSE _State = TEST_RUN_PHASE.REPORTING_TOTALS THEN
	RETURN;
END_IF

IF ExitCode = -1 THEN
	validateChildren(rejectRunningChildren := FALSE);

	FOR i := 0 TO _ChildCount - 1 DO
		Children[i].Reset(reporter := 0);
	END_FOR
END_IF

TOF_Core.DynamicMemoryManager.RaiseIfAllocationFailed();

IsFinished := FALSE;
AllPassed := FALSE;
ExitCode := 0;
CallbackException := __SYSTEM.ExceptionCode.RTSEXCPT_NOEXCEPTION;
CallbackMessage := "";
TotalTests := 0;
PassedTests := 0;
FailedTests := 0;
SkippedTests := 0;
TotalDuration := T#0S;

_State := TEST_RUN_PHASE.STARTING;
_CurrentChildIndex := 0;
_Duration := LTIME#0NS;
END_METHOD

(*!
<summary>Checks the fixed root array before startup or explicit abort recovery.</summary>
<description>
Missing storage or null slots raise DataMemberNotSpecifiedException; duplicate or group-owned roots raise
StandardException. Startup also rejects running roots. Abort recovery permits running roots so their Reset
callbacks can recover execution state after the caller has made user resources safe. Failures propagate
without calling any child or changing runner observations. No allocation occurs for a valid composition.
</description>
<param name="rejectRunningChildren">TRUE for startup; FALSE for explicit recovery of an aborted tree.</param>
*)
METHOD PRIVATE validateChildren
VAR_INPUT
	rejectRunningChildren : BOOL;
END_VAR
VAR
	i : INT;
	j : INT;
	childParent : ITestElement;
	
	errorMessage : TOF_Core.ERROR_MESSAGE;
END_VAR
IF NOT __ISVALIDREF(Children) THEN
	TOF_Core.Exceptions.ThrowDataMemberNotSpecified(
		sourceNamespaceName := NamespaceName,
		sourceClassName := ClassName,
		sourcePOUName := __POUNAME(),
		sourcePosition := __POSITION(),
		dataMemberName := 'Children'
	);
END_IF

FOR i := 0 TO _ChildCount - 1 DO
	IF Children[i] = 0 THEN
		TOF_Core.Exceptions.ThrowDataMemberNotSpecified(
			sourceNamespaceName := NamespaceName,
			sourceClassName := ClassName,
			sourcePOUName := __POUNAME(),
			sourcePosition := __POSITION(),
			dataMemberName := TOF_Core.Strings.Concat255('Children[', TO_STRING(i), ']')
		);
	END_IF

	childParent := Children[i].Parent;

	IF childParent <> 0 THEN
		errorMessage := TOF_Core.WideStrings.Concat255("A root child '", Children[i].Name, "' belongs to a group");

		TOF_Core.Exceptions.ThrowStandard(
			sourceNamespaceName := NamespaceName,
			sourceClassName := ClassName,
			sourcePOUName := __POUNAME(),
			sourcePosition := __POSITION(),
			message := errorMessage
		);
	END_IF

	IF rejectRunningChildren AND_THEN Children[i].IsRunning THEN
		errorMessage := TOF_Core.WideStrings.Concat255("A root child '", Children[i].Name, "' is active");
 
		TOF_Core.Exceptions.ThrowStandard(
			sourceNamespaceName := NamespaceName,
			sourceClassName := ClassName,
			sourcePOUName := __POUNAME(),
			sourcePosition := __POSITION(),
			message := errorMessage
		);
	END_IF

	FOR j := 0 TO i - 1 DO
		IF Children[i] = Children[j] THEN
			errorMessage := TOF_Core.WideStrings.Concat255("A root child '", Children[i].Name, "' occupies more than one slot"); 
			
			TOF_Core.Exceptions.ThrowStandard(
				sourceNamespaceName := NamespaceName,
				sourceClassName := ClassName,
				sourcePOUName := __POUNAME(),
				sourcePosition := __POSITION(),
				message := errorMessage
			);
		END_IF
	END_FOR
END_FOR
END_METHOD

END_FUNCTION_BLOCK

// ---- TestElements/Tests/SingleCycleTest.TcPOU
(*
SPDX-FileCopyrightText: © 2026 Oleksandr Tiutyk <trofimich@gmail.com>
SPDX-License-Identifier: MIT
License: https://opensource.org/license/mit
*)

(*!
<summary>Base class for one test whose body completes in a single PLC scheduling cycle.</summary>
<description>
Override ExecuteTest with the checks. Returning from the body completes the body automatically.
BeforeTest and AfterTest are optional scenario hooks. Constructor name identifies the case in reports.
Run through TestRunner, directly or inside a TestGroup. A complete run and its reporting may span more cycles
than the body. All instance access belongs to one task without reentry; other tasks need other instances.
</description>
*)

{attribute 'no_explicit_call' := 'do not call this function block directly'}
FUNCTION_BLOCK ABSTRACT SingleCycleTest EXTENDS TestCase

(*!
<summary>Implements the scenario body without runner guards or enumeration.</summary>
<description>
Keep persistent state in instance fields. Reporting a failure does not abort the current callback.
</description>
*)
METHOD PROTECTED ABSTRACT ExecuteTest
END_METHOD

(*!
<summary>Runs the body once and reports completion for the cycle.</summary>
*)
METHOD PROTECTED FINAL RunCycle : TEST_CYCLE_RESULT
ExecuteTest();
RunCycle := TEST_CYCLE_RESULT.DONE;
END_METHOD

END_FUNCTION_BLOCK

// ---- TestElements/Tests/MultiCycleTest.TcPOU
(*
SPDX-FileCopyrightText: © 2026 Oleksandr Tiutyk <trofimich@gmail.com>
SPDX-License-Identifier: MIT
License: https://opensource.org/license/mit
*)

(*!
<summary>Base class for one test that waits or advances state across PLC scheduling cycles.</summary>
<description>
Override ExecuteTest with one bounded step returning TEST_CYCLE_RESULT.BUSY to await the next task cycle or
TEST_CYCLE_RESULT.DONE when finished. BeforeTest prepares once and AfterTest cleans up once, including failure.
Timeout defaults to one second; zero disables it. A nonzero deadline is checked before every body after the first.
Once a cycle returns DONE and finishes the case, subsequent cycles do not run. Timing sums nominal task periods,
not wall-clock time. Use a typed enumeration in the derived FB when the scenario needs a state machine. No numeric
step API is used. Each instance belongs to one task without reentry. Constructor name identifies the case in reports.
</description>
*)

{attribute 'no_explicit_call' := 'do not call this function block directly'}
FUNCTION_BLOCK ABSTRACT MultiCycleTest EXTENDS TestCase
VAR
	_Timeout : TIME := T#1S;
END_VAR

(*!
<summary>Implements one bounded scenario step and reports whether execution continues or is done.</summary>
<description>
Keep persistent state in instance fields. Return TEST_CYCLE_RESULT.BUSY to wait for the next task cycle or
TEST_CYCLE_RESULT.DONE when finished. Reporting a failure does not abort the current callback, and any failure
terminates the case after the callback returns even if BUSY is returned.
</description>
*)
METHOD PROTECTED ABSTRACT ExecuteTest : TEST_CYCLE_RESULT
END_METHOD

(*!
<summary>Checks the deadline before advancing one body cycle.</summary>
*)
METHOD PROTECTED FINAL RunCycle : TEST_CYCLE_RESULT
IF _Timeout > T#0S AND_THEN _Elapsed >= TO_LTIME(_Timeout) THEN
	RecordFailure(message := "Multi-cycle test exceeded deadline");
	RunCycle := TEST_CYCLE_RESULT.DONE;
ELSE
	RunCycle := ExecuteTest();
END_IF
END_METHOD

(*!
<summary>Gets or configures the whole-scenario deadline; zero disables it.</summary>
<description>
Configure before execution or after completion. Mutation during a run raises StandardException
because the operation is invalid in the current state, regardless of the requested deadline value.
</description>
*)
{attribute 'monitoring' := 'call'}
PROPERTY Timeout : TIME
GET
Timeout := _Timeout;
END_GET
SET
IF IsRunning THEN
	TOF_Core.Exceptions.ThrowStandard(
		sourceNamespaceName := NamespaceName,
		sourceClassName := ClassName,
		sourcePOUName := __POUNAME(),
		sourcePosition := __POSITION(),
		message := "Cannot change an active test deadline"
	);
END_IF

_Timeout := Timeout;
END_SET
END_PROPERTY

END_FUNCTION_BLOCK
